TYPE ST_Interlock :
STRUCT
	conditions	: ARRAY[1..10] OF BOOL := [1,1,1,1,1,1,1,1,1,1];
	descriptions	: ARRAY[1..10] OF STRING := ['N/A','N/A','N/A','N/A','N/A','N/A','N/A','N/A','N/A','N/A'];
END_STRUCT
END_TYPE

(* stored: Version 1.1.0.1
   DUT ST_Interlock: Id {4300dd3d-cb05-43eb-a93d-e40bc8ef5461} *)
